{attribute 'no_assign'}
FUNCTION_BLOCK FB_LD_WTURBINELD0 EXTENDS FB_AcsiCommonLogicalDeviceClass
VAR_INPUT
	LLN0: FB_LN_WTURBINE_LD0_LLN0 := (sClass:='LLN0', bLinkResult:=THIS^.AddLogicalNodeToContainer(ipLogicalNode:=LLN0));
	LPHD1: FB_LN_WTURBINE_LD0_LPHD1 := (sClass:='LPHD', bLinkResult:=THIS^.AddLogicalNodeToContainer(ipLogicalNode:=LPHD1));
	WGEN1: FB_LN_WTURBINE_LD0_WGEN1 := (sClass:='WGEN', bLinkResult:=THIS^.AddLogicalNodeToContainer(ipLogicalNode:=WGEN1));
	WTUR1: FB_LN_WTURBINE_LD0_WTUR1 := (sClass:='WTUR', bLinkResult:=THIS^.AddLogicalNodeToContainer(ipLogicalNode:=WTUR1));
	WROT1: FB_LN_WTURBINE_LD0_WROT1 := (sClass:='WROT', bLinkResult:=THIS^.AddLogicalNodeToContainer(ipLogicalNode:=WROT1));
	WCNV1: FB_LN_WTURBINE_LD0_WCNV1 := (sClass:='WCNV', bLinkResult:=THIS^.AddLogicalNodeToContainer(ipLogicalNode:=WCNV1));
	WMET1: FB_LN_WTURBINE_LD0_WMET1 := (sClass:='WMET', bLinkResult:=THIS^.AddLogicalNodeToContainer(ipLogicalNode:=WMET1));
	WALM1: FB_LN_WTURBINE_LD0_WALM1 := (sClass:='WALM', bLinkResult:=THIS^.AddLogicalNodeToContainer(ipLogicalNode:=WALM1));
	WYAW1: FB_LN_WTURBINE_LD0_WYAW1 := (sClass:='WYAW', bLinkResult:=THIS^.AddLogicalNodeToContainer(ipLogicalNode:=WYAW1));
	WPPD1: FB_LN_WTURBINE_LD0_WPPD1 := (sClass:='WPPD', bLinkResult:=THIS^.AddLogicalNodeToContainer(ipLogicalNode:=WPPD1));
END_VAR
VAR
END_VAR

END_FUNCTION_BLOCK

(* stored: Version 1.1.0.1
   POU FB_LD_WTURBINELD0: Id {1fe18e34-e772-4cbd-a9d9-75a8dcceb6e6}, SpecialFunc None *)
